FUNCTION_BLOCK ProjectInformation_Tests EXTENDS TcUnit.FB_TestSuite

Test_VersionIsFourPointTwo();
Test_TitleAndCompany();

METHOD PRIVATE Test_VersionIsFourPointTwo
VAR
  version : ST_LibVersion;
END_VAR
TcUnit.TEST(__POUNAME());

version := F_GetVersion();
AssertEquals_STRING(Expected := '4.2.0.0', Actual := version.sVersion, Message := 'library version string');
AssertEquals_UINT(Expected := 4, Actual := version.iMajor, Message := 'major version');
AssertEquals_UINT(Expected := 2, Actual := version.iMinor, Message := 'minor version');

TEST_FINISHED_NAMED(__POUNAME());
END_METHOD

METHOD PRIVATE Test_TitleAndCompany
TcUnit.TEST(__POUNAME());

AssertEquals_WSTRING(Expected := "Intecre.Utilities", Actual := F_GetTitle(), Message := 'library title');
AssertEquals_WSTRING(Expected := "Intecre Ltd", Actual := F_GetCompany(), Message := 'library company');

TEST_FINISHED_NAMED(__POUNAME());
END_METHOD

END_FUNCTION_BLOCK

(* stored: Version 1.1.0.1, ProductVersion 3.1.4026.22
   POU ProjectInformation_Tests: Id {6c643318-cb51-463a-86cd-2b298e83f5d7}, SpecialFunc None
   Method Test_VersionIsFourPointTwo: Id {a479a1da-6388-4562-8a17-5e0761ca0380}
   Method Test_TitleAndCompany: Id {9533a47f-f557-4686-b84c-a1c50544af0e} *)
